Fanuc KAREL source: KT00877.KL

PROGRAM KT00877
%NOLOCKGROUP
VAR
  B1: BOOLEAN
  B2: BOOLEAN
  OUT: REAL
BEGIN
  B1 = TRUE
  B2 = FALSE
  B1 = TRUE
  B2 = FALSE
  OUT = TRUNC(B1)
END KT00877
